Staubli VAL3: teachPoint.pgx

program teachPoint(num x_nStep, num x_nIndex)
  local bool l_bResult
begin
  l_bResult=userPageConfirm("是否记录该点位？")
  if l_bResult
    switch x_nStep
      case 0
        savedata:fFrameItem[x_nIndex].pPointRx[0]=here(tUsingTool,world)
      break
      case 1
        savedata:fFrameItem[x_nIndex].pPointRx[1]=here(tUsingTool,world)
      break
      case 2
        savedata:fFrameItem[x_nIndex].pPointRx[2]=here(tUsingTool,world)
      break

    endSwitch
  endIf
end
